Staubli VAL3: onStart.pgx

public program onStart()
  local num l_nSize
  local string l_sMsg
  local num l_i
begin
  sLstValue=""
  nPageIndex=0
  nPageNum=1
  call refreshlist()

  sPageIndex=toString("",nPageIndex+1)
  sPageNum=toString("",nPageNum)
end
